(*
SPDX-FileCopyrightText: © 2026 Oleksandr Tiutyk <trofimich@gmail.com>
SPDX-License-Identifier: MIT
License: https://opensource.org/license/mit
*)

(*!
<summary>Exposes the object's current error status and diagnostic details.</summary>
<description>
Error storage belongs to the provider. Changes and clearing follow the provider's lifecycle.
</description>
*)

INTERFACE IErrorProvider EXTENDS IObject

(*!
<summary>Returns a borrowed, read-only view of the current diagnostic error.</summary>
<description>
Callers must not modify fields or call mutating methods such as Clear or SetSeverity through this reference.
The view requires a live provider and may change when the provider updates its error state.
</description>
*)

{attribute 'monitoring' := 'call'}
PROPERTY Error : REFERENCE TO ERROR
GET
END_GET
END_PROPERTY

(*!
<summary>Reports whether the current Error represents an error.</summary>
<description>
This is the provider's current status, not an indication that its operation has completed.
</description>
*)

{attribute 'monitoring' := 'call'}
PROPERTY HasError : BOOL
GET
END_GET
END_PROPERTY

END_INTERFACE

(* stored: Version 1.1.0.1
   Itf IErrorProvider: Id {5f0d4ebb-811f-4762-ade5-09da7d3b686c}
   Property Error: Id {a23ffa71-c915-4bac-a195-e5f5c3765f25}
   Get Get: Id {06944b97-05cd-462c-b84e-f1632ad8c537}
   Property HasError: Id {2988e528-f3cf-437a-ad0d-0bd717afcf95}
   Get Get: Id {a5906d11-aa99-468b-928a-9e1895366cbe} *)
